// TIA Portal V20 export
// export: Created 2026-10-20T12:52:50.1330528Z, ExportSetting WithDefaults, DisplayName Totally Integrated Automation Portal, DisplayVersion V20 Update 6, DisplayName TIA Portal Openness, DisplayVersion V20 Update 6, DisplayName TIA Portal Version Control Interface, DisplayVersion V20 Update 6, DisplayName SINAMICS Startdrive Advanced, DisplayVersion V20 SP1, DisplayName SINAMICS Startdrive G130, G150, S120, S150, SINAMICS MV, G220, S200, S210, DisplayVersion V20 SP1, DisplayName SINAMICS Startdrive G110M, G120, G120C, G120D, G120P, G115D, DisplayVersion V20 SP1, DisplayName STEP 7 Professional, DisplayVersion V20 Update 6, DisplayName STEP 7 Safety, DisplayVersion V20 Update 2, DisplayName WinCC Basic/Comfort/Advanced, DisplayVersion V20 Update 6, DisplayName WinCC Unified, DisplayVersion V20 Update 6
FUNCTION "Handshake_Outfeed_FC" : Void   // FC51, SCL
{ S7_Optimized_Access := 'TRUE' }
VERSION : 0.1
// stored: AutoNumber true, IsIECCheckEnabled false, SetENOAutomatically false, UDAEnableTagReadback false
   VAR_INPUT
      Auto_Mode : Bool;
      Ready_To_Send : Bool;
      Conv_Occupied : Bool;
      Transfer_In_Progress : Bool;
      DB_LGX_To_SM_Outfeed_Ready_To_Receive : Bool;
   END_VAR
   VAR_OUTPUT
      Fault_Handshake : Bool;
      DB_SM_To_LGX_Outfeed_Transfer_In_Progress : Bool;
      DB_SM_To_LGX_Outfeed_Ocuppied : Bool;
      DB_SM_To_LGX_Outfeed_Ready_To_Send : Bool;
   END_VAR
   VAR_TEMP
      tCanSend : Bool;
   END_VAR
BEGIN
   // ---------------------------------------------------------
   // STEP 1: Is SM ready to send?
   // Condition: pallet waiting at exit, SM in auto,
   //            no transfer in progress
   // ---------------------------------------------------------
   #tCanSend :=
   #Auto_Mode
   AND #Conv_Occupied
   AND #Ready_To_Send
   AND NOT #DB_SM_To_LGX_Outfeed_Transfer_In_Progress;

   IF #tCanSend
       AND NOT #DB_SM_To_LGX_Outfeed_Ready_To_Send THEN
       #DB_SM_To_LGX_Outfeed_Ready_To_Send := TRUE;
   END_IF;

   // ---------------------------------------------------------
   // STEP 2: LGX responded Ready_To_Receive → start transfer
   // ---------------------------------------------------------
   IF NOT #Conv_Occupied THEN
       // #DB_SM_To_LGX_Outfeed_Transfer_In_Progress := TRUE;
       #DB_SM_To_LGX_Outfeed_Ready_To_Send := FALSE;
   END_IF;

   // ---------------------------------------------------------
   // STEP 3: LGX confirmed pallet received
   // → SM resets Transfer_In_Progress
   // ---------------------------------------------------------
   // IF #DB_SM_To_LGX_Outfeed_Transfer_In_Progress
   //     AND #DB_LGX_To_SM_Outfeed_Ready_To_Receive THEN
   //     #DB_SM_To_LGX_Outfeed_Transfer_In_Progress := FALSE;
   // END_IF;

   #DB_SM_To_LGX_Outfeed_Transfer_In_Progress := #Transfer_In_Progress;
   #DB_SM_To_LGX_Outfeed_Ocuppied := #Conv_Occupied;
   // ---------------------------------------------------------
   // STEP 4: Reset Ready_To_Send if pallet removed or SM left auto mode
   // ---------------------------------------------------------
   IF NOT #Ready_To_Send OR NOT #Auto_Mode THEN
       IF NOT #DB_SM_To_LGX_Outfeed_Transfer_In_Progress THEN
           #DB_SM_To_LGX_Outfeed_Ready_To_Send := FALSE;
       END_IF;
   END_IF;

   #Fault_Handshake := FALSE; // Placeholder
END_FUNCTION
